TYPE ST_WorkshopOutputs :
STRUCT
    bLightRelay : BOOL;
END_STRUCT
END_TYPE

(* stored: Version 1.1.0.1
   DUT ST_WorkshopOutputs: Id {c193ec37-15dd-46b0-914a-80dcdd01fd86} *)
